(* IEC 61131-3 sources: codesys-to-s7/tests/corpus/C2S7-TYPE-TIME/neg, 1 file *)

(* ---- input.st ---- *)
FUNCTION_BLOCK FB_Case
VAR
    a : INT;
    b : INT;
    i : INT;
    d : DINT;
    r : REAL;
    x : BOOL;
    y : BOOL;
    s : STRING(80);
    w : WORD;
    t : TIME;
END_VAR
t := T#10D;
END_FUNCTION_BLOCK
